SUBAPPLICATION mapping_Buttons (* Subapplication Type *)
  (* Standard: 61499-2 *)
  (* Version 1.0, 2023-01-29, Franz *)
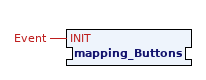
  EVENT_INPUT
    INIT;
  END_EVENT
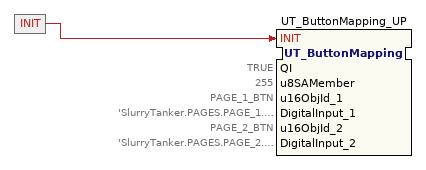
  FBS
    UT_ButtonMapping_UP : UT_ButtonMapping(QI := TRUE, u8SAMember := 255, u16ObjId_1 := PAGE_1_BTN, DigitalInput_1 := 'SlurryTanker.PAGES.PAGE_1.BTN', u16ObjId_2 := PAGE_2_BTN, DigitalInput_2 := 'SlurryTanker.PAGES.PAGE_2.BTN');
  END_FBS
  EVENT_CONNECTIONS
    INIT TO UT_ButtonMapping_UP.INIT;
  END_CONNECTIONS
END_SUBAPPLICATION
